        bool bMouseDown
        bool bMouseUp
    utText Text
      [0]
        num nFontSize
        string sFontFamily
        string sFontStyle
        string sFontWeight
        string sTextAlignment
public utLabel utLbl_Tool
  [0]
    utAppearance Appearance
      [0]
        bool bVisibility
        string sBackgroundColour = "#FFFFFF"
        string sColour
    utBorder Border
      [0]
        num nBorderWidth
        string sBorderColour
        string sBorderStyle
    utCommon Common
      [0]
        string sID = "lbl_Tool"
        string sPage = "Disk://SmartTCP_CS9/ts2/interface/Page_Main"
        string sText = "工具："
    utData Data
      [0]
        bool bStatus
        num nVal = 99
    utEvents Events
      [0]
        bool bClick
        bool bMouseDown
        bool bMouseUp
    utText Text
      [0]
        num nFontSize
        string sFontFamily
        string sFontStyle
        string sFontWeight
        string sTextAlignment
public utLabel utLbl_ToolValue_Data[6]
  [0]
    utAppearance Appearance
      [0]
        bool bVisibility
        string sBackgroundColour = "#FFFFFF"
        string sColour
    utBorder Border
      [0]
        num nBorderWidth
        string sBorderColour
        string sBorderStyle
    utCommon Common
      [0]
        string sID = "utLbl_ToolValue_Data0"
        string sPage = "Disk://SmartTCP_CS9/ts2/interface/Page_Container_Test"
        string sText = "120    "
    utData Data
      [0]
        bool bStatus
        num nVal = 99
    utEvents Events
      [0]
        bool bClick
        bool bMouseDown
        bool bMouseUp
    utText Text
      [0]
        num nFontSize
        string sFontFamily
        string sFontStyle
        string sFontWeight
        string sTextAlignment
  [1]
    utAppearance Appearance
      [0]
        bool bVisibility
        string sBackgroundColour = "#FFFFFF"
        string sColour
    utBorder Border
      [0]
        num nBorderWidth
        string sBorderColour
        string sBorderStyle
    utCommon Common
      [0]
        string sID = "utLbl_ToolValue_Data1"
        string sPage = "Disk://SmartTCP_CS9/ts2/interface/Page_Container_Test"
        string sText = "55    "
    utData Data
      [0]
        bool bStatus
        num nVal = 99
    utEvents Events
      [0]
        bool bClick
        bool bMouseDown
        bool bMouseUp
    utText Text
      [0]
        num nFontSize
        string sFontFamily
        string sFontStyle
        string sFontWeight
        string sTextAlignment
  [2]
    utAppearance Appearance
      [0]
        bool bVisibility
        string sBackgroundColour = "#FFFFFF"
        string sColour
    utBorder Border
      [0]
        num nBorderWidth
        string sBorderColour
        string sBorderStyle
    utCommon Common
      [0]
        string sID = "utLbl_ToolValue_Data2"
        string sPage = "Disk://SmartTCP_CS9/ts2/interface/Page_Container_Test"
        string sText = "0    "
    utData Data
      [0]
        bool bStatus
        num nVal = 99
    utEvents Events
      [0]
        bool bClick
        bool bMouseDown
        bool bMouseUp
    utText Text
      [0]
        num nFontSize
        string sFontFamily
        string sFontStyle
        string sFontWeight
        string sTextAlignment
  [3]
    utAppearance Appearance
      [0]
        bool bVisibility
        string sBackgroundColour = "#FFFFFF"
        string sColour
    utBorder Border
      [0]
        num nBorderWidth
        string sBorderColour
        string sBorderStyle
    utCommon Common
      [0]
        string sID = "utLbl_ToolValue_Data3"
        string sPage = "Disk://SmartTCP_CS9/ts2/interface/Page_Container_Test"
        string sText = "0    "
    utData Data
      [0]
        bool bStatus
        num nVal = 99
    utEvents Events
      [0]
        bool bClick
        bool bMouseDown
        bool bMouseUp
    utText Text
      [0]
        num nFontSize
        string sFontFamily
        string sFontStyle
        string sFontWeight
        string sTextAlignment
  [4]
    utAppearance Appearance
      [0]
        bool bVisibility
        string sBackgroundColour = "#FFFFFF"
        string sColour
    utBorder Border
      [0]
        num nBorderWidth
        string sBorderColour
        string sBorderStyle
    utCommon Common
      [0]
        string sID = "utLbl_ToolValue_Data4"
        string sPage = "Disk://SmartTCP_CS9/ts2/interface/Page_Container_Test"
        string sText = "0    "
    utData Data
      [0]
        bool bStatus
        num nVal = 99
    utEvents Events
      [0]
        bool bClick
        bool bMouseDown
        bool bMouseUp
    utText Text
      [0]
        num nFontSize
        string sFontFamily
        string sFontStyle
        string sFontWeight
        string sTextAlignment
  [5]
    utAppearance Appearance
      [0]
        bool bVisibility
        string sBackgroundColour = "#FFFFFF"
        string sColour
    utBorder Border
      [0]
        num nBorderWidth
        string sBorderColour
        string sBorderStyle
    utCommon Common
      [0]
        string sID = "utLbl_ToolValue_Data5"
        string sPage = "Disk://SmartTCP_CS9/ts2/interface/Page_Container_Test"
        string sText = "0    "
    utData Data
      [0]
        bool bStatus
        num nVal = 99
    utEvents Events
      [0]
        bool bClick
        bool bMouseDown
        bool bMouseUp
    utText Text
      [0]
        num nFontSize
        string sFontFamily
        string sFontStyle
        string sFontWeight
        string sTextAlignment
public utLabel utLbl_Tool_Data
  [0]
    utAppearance Appearance
      [0]
        bool bVisibility
        string sBackgroundColour = "#FFFFFF"
        string sColour
    utBorder Border
      [0]
        num nBorderWidth
        string sBorderColour
        string sBorderStyle
    utCommon Common
      [0]
        string sID = "lbl_Tool_Data"
        string sPage = "Disk://SmartTCP_CS9/ts2/interface/Page_Main"
        string sText = "tFlange"
    utData Data
      [0]
        bool bStatus
        num nVal = 99
    utEvents Events
      [0]
        bool bClick
        bool bMouseDown
        bool bMouseUp
    utText Text
      [0]
        num nFontSize
        string sFontFamily
        string sFontStyle
        string sFontWeight
        string sTextAlignment
public utText utTxt_OffsetValue_Data[6]
  [0]
    utAppearance Appearance
      [0]
        bool bVisibility
        string sBackgroundColour = "#EEFF00"
        string sColour
    utBorder Border
      [0]
        string sBorderColour
        string sBorderSytle
        string sBorderWidth
    utCommon Common
      [0]
        bool bDisabled
        num nValue
        string sID = "utTxt_OffsetValue_Data0"
        string sPage = "Disk://SmartTCP_CS9/ts2/interface/Page_Container_Test"
        string sValue
    utText Text
      [0]
        num nFontSize
        string sFontFamily
        string sFontStyle
        string sFontWeight
        string sTextAlignment
  [1]
    utAppearance Appearance
      [0]
        bool bVisibility
        string sBackgroundColour = "#EEFF00"
        string sColour
    utBorder Border
      [0]
        string sBorderColour
        string sBorderSytle
        string sBorderWidth
    utCommon Common
      [0]
        bool bDisabled
        num nValue
        string sID = "utTxt_OffsetValue_Data1"
        string sPage = "Disk://SmartTCP_CS9/ts2/interface/Page_Container_Test"
        string sValue
    utText Text
      [0]
        num nFontSize
        string sFontFamily
        string sFontStyle
        string sFontWeight
        string sTextAlignment
  [2]
    utAppearance Appearance
      [0]
        bool bVisibility
        string sBackgroundColour = "#EEFF00"
        string sColour
    utBorder Border
      [0]
        string sBorderColour
        string sBorderSytle
        string sBorderWidth
    utCommon Common
      [0]
        bool bDisabled
        num nValue = 10
        string sID = "utTxt_OffsetValue_Data2"
        string sPage = "Disk://SmartTCP_CS9/ts2/interface/Page_Container_Test"
        string sValue
    utText Text
      [0]
        num nFontSize
        string sFontFamily
        string sFontStyle
        string sFontWeight
        string sTextAlignment
  [3]
    utAppearance Appearance
      [0]
        bool bVisibility
        string sBackgroundColour = "#EEFF00"
        string sColour
    utBorder Border
      [0]
        string sBorderColour
        string sBorderSytle
        string sBorderWidth
    utCommon Common
      [0]
        bool bDisabled
        num nValue
        string sID = "utTxt_OffsetValue_Data3"
        string sPage = "Disk://SmartTCP_CS9/ts2/interface/Page_Container_Test"
        string sValue
    utText Text
      [0]
        num nFontSize
        string sFontFamily
        string sFontStyle
        string sFontWeight
        string sTextAlignment
  [4]
    utAppearance Appearance
      [0]
        bool bVisibility
        string sBackgroundColour = "#EEFF00"
        string sColour
    utBorder Border
      [0]
        string sBorderColour
        string sBorderSytle
        string sBorderWidth
    utCommon Common
      [0]
        bool bDisabled
        num nValue
        string sID = "utTxt_OffsetValue_Data4"
        string sPage = "Disk://SmartTCP_CS9/ts2/interface/Page_Container_Test"
        string sValue
    utText Text
      [0]
        num nFontSize
        string sFontFamily
        string sFontStyle
        string sFontWeight
        string sTextAlignment
  [5]
    utAppearance Appearance
      [0]
        bool bVisibility
        string sBackgroundColour = "#EEFF00"
        string sColour
    utBorder Border
      [0]
        string sBorderColour
        string sBorderSytle
        string sBorderWidth
    utCommon Common
      [0]
        bool bDisabled
        num nValue
        string sID = "utTxt_OffsetValue_Data5"
        string sPage = "Disk://SmartTCP_CS9/ts2/interface/Page_Container_Test"
        string sValue
    utText Text
      [0]
        num nFontSize
        string sFontFamily
        string sFontStyle
        string sFontWeight
        string sTextAlignment
public utText utTxt_popUpMsg
  [0]
    utAppearance Appearance
      [0]
        bool bVisibility
        string sBackgroundColour = "#7C95FF"
        string sColour
    utBorder Border
      [0]
        string sBorderColour
        string sBorderSytle
        string sBorderWidth
    utCommon Common
      [0]
        bool bDisabled
        num nValue
        string sID = "txt_popUpMsg"
        string sPage = "Disk://SmartTCP_CS9/ts2/interface/Page_Container_Confirm"
        string sValue = "第2点记录完成"
    utText Text
      [0]
        num nFontSize
        string sFontFamily
        string sFontStyle
        string sFontWeight
        string sTextAlignment
public utTool utCurrentTool
  [0]
    num nItem
    num nItemM = 1
    string sName
    tool tValue = {fatherId=flange[0]}
